Staubli VAL3: _clickProductionPage.pgx

public program _clickProductionPage()
begin
  sPageUsing="cycleCtrl"
  userPage("Disk://Project/interface/cycleCtrl")
  delay(1)
end
